// TIA Portal V20 export
Screen "Screen_1"  1366x768
